Fanuc KAREL source: KD00042.KL

PROGRAM KD00042
%NOLOCKGROUP
VAR
  I: INTEGER
  J: INTEGER
  B: BOOLEAN
  R: REAL
  S: STRING[80]
  N: STD_PTH_NODE
BEGIN
  I = 1
END KD00042
